(* IEC 61131-3 sources: st2fb/corpus_hard/public_st/p01_bistable_device, 2 files *)

(* ---- control_flat.st ---- *)
(* Solvability control, never shown to a model: the same behaviour in the translator's v1 subset, written for this project.
   The only change is that USINT became INT, and input initial values were dropped since the harness writes every input. *)
FUNCTION_BLOCK GenericBistableDeviceModel
VAR_INPUT
  ActivateCmd : BOOL;
  DeactivateCmd : BOOL;
  cfgActTime : TIME;
  cfgDeactTime : TIME;
  simActFail : BOOL;
  simDeactFail : BOOL;
END_VAR
VAR_OUTPUT
  Activated : BOOL;
  Deactivated : BOOL;
END_VAR
VAR
  TransitionDelay : TON;
  vState : INT := 0;
  vStateOld : INT := 3;
END_VAR
CASE vState OF
  0:
    IF vState <> vStateOld THEN
      TransitionDelay(IN := FALSE);
      vStateOld := vState;
    END_IF;
    TransitionDelay(IN := ActivateCmd AND NOT simActFail, PT := cfgActTime);
    IF TransitionDelay.Q THEN
      vState := 1;
    END_IF;
  1:
    IF vState <> vStateOld THEN
      TransitionDelay(IN := FALSE);
      vStateOld := vState;
    END_IF;
    TransitionDelay(IN := DeactivateCmd AND NOT simDeactFail, PT := cfgDeactTime);
    IF TransitionDelay.Q THEN
      vState := 0;
    END_IF;
END_CASE;
Activated := vState = 1;
Deactivated := vState = 0;
END_FUNCTION_BLOCK

(* ---- program.st ---- *)
(* From tkucic/plc_hello_mixing_tank, GenericBistableDeviceModel. Copyright (c) 2021 Toni Kucic. MIT licence, see LICENSE
   in this directory. *)
FUNCTION_BLOCK GenericBistableDeviceModel
VAR_INPUT
  ActivateCmd : BOOL;
  DeactivateCmd : BOOL;
  cfgActTime : TIME := TIME#1s0ms;
  cfgDeactTime : TIME := TIME#1s0ms;
  simActFail : BOOL;
  simDeactFail : BOOL;
END_VAR
VAR_OUTPUT
  Activated : BOOL;
  Deactivated : BOOL;
END_VAR
VAR
  TransitionDelay : TON;
  vState : USINT := 0;
  vStateOld : USINT := 3;
END_VAR
CASE vState OF
	0: (*Deactivated*)
		(*On entry do:*)
		IF vState <> vStateOld THEN
			(*Reset timer*)
			TransitionDelay(IN:=FALSE);
			vStateOld := vState;
		END_IF;
		TransitionDelay(IN:=ActivateCmd AND NOT simActFail, PT:=cfgActTime);
		IF TransitionDelay.Q THEN
			vState := 1;
		END_IF;
	1: (*Activated*)
		(*On entry do:*)
		IF vState <> vStateOld THEN
			(*Reset timer*)
			TransitionDelay(IN:=FALSE);
			vStateOld := vState;
		END_IF;
		TransitionDelay(IN:=DeactivateCmd AND NOT simDeactFail, PT:=cfgDeactTime);
		IF TransitionDelay.Q THEN
			vState := 0;
		END_IF;
END_CASE;
Activated := vState = 1;
Deactivated := vState = 0;
END_FUNCTION_BLOCK
